(* IEC 61131-3 sources: PLC-Static-Analysis/modules/plc-rules/src/test/resources/PLCA-L024, 2 files *)

(* ---- compliant.st ---- *)
PROGRAM P_L024ok
VAR
    n : INT;
    m : INT;
    r : REAL;
    b : BOOL;
    c : BOOL;
    q : BOOL;
END_VAR
q := n <> 10;
q := NOT b;
q := NOT (b AND c);
END_PROGRAM

(* ---- noncompliant.st ---- *)
PROGRAM P_L024
VAR
    n : INT;
    m : INT;
    r : REAL;
    b : BOOL;
    c : BOOL;
    q : BOOL;
END_VAR
q := NOT (n = 10); // PLCA-L024
IF NOT (n < m) THEN // PLCA-L024
    q := TRUE;
END_IF
END_PROGRAM
